Staubli VAL3: HMI_util.pjx

--- HMI_util.pjx ---
Parameters version=s8.12.2Cs9_BS2561 stackSize=5000 millimeterUnit=true
Program file=initJogMode.pgx
Program file=jogMode.pgx
Program file=loadingPage.pgx
Program file=login.pgx
Program file=setBtnColor.pgx
Program file=setframemode.pgx
Program file=setjointmode.pgx
Program file=setnullmode.pgx
Program file=settoolmode.pgx
Program file=start.pgx
Program file=stop.pgx
Data file=HMI_util.dtx
Library alias=savedata path=Disk://source/saveData/saveData.pjx

--- HMI_util.dtx ---
mdesc mNomSpeed
public string sShowType[6]
public string sShowNum[6]
public string sJoint[6]
  [0] = "J1:"
  [1] = "J2:"
  [2] = "J3:"
  [3] = "J4:"
  [4] = "J5:"
  [5] = "J6:"
public string sCartisiam[6]
  [0] = "X:"
  [1] = "Y:"
  [2] = "Z:"
  [3] = "RX:"
  [4] = "RY:"
  [5] = "RZ:"
public string sPage
string sInputPswd
bool bConfirm
bool bCancel
string sPassword = "1"
num nUsingTool

--- start.pgx ---
program start()
begin
end

--- initJogMode.pgx ---
public program initJogMode()
  local num l_i
begin
   for l_i = 0 to size(sShowType)-1
    sShowType[l_i]=sCartisiam[l_i]
  endFor
end

--- jogMode.pgx ---
public program jogMode(num x_nToolIndex, num x_nFrameIndex)
  local num l_nJogMode
  local jointRx l_jHere
  local pointRx l_pHere
  local tool l_tTool
  local frame l_fFrame
begin
  link(l_tTool,flange)
  link(l_fFrame,world)
  l_nJogMode=$getJogmode()
  l_jHere=herej()
  call savedata:getTool(x_nToolIndex,l_tTool)
  call savedata:getFrame(x_nFrameIndex,l_fFrame)
  l_pHere=here(l_tTool,l_fFrame)
  switch l_nJogMode
    case 0
      call setBtnColor(0)
      sShowNum[0]=toString(".2",l_pHere.trsf.x)
      sShowNum[1]=toString(".2",l_pHere.trsf.y)
      sShowNum[2]=toString(".2",l_pHere.trsf.z)
      sShowNum[3]=toString(".2",l_pHere.trsf.rx)
      sShowNum[4]=toString(".2",l_pHere.trsf.ry)
      sShowNum[5]=toString(".2",l_pHere.trsf.rz )
    break
    case 1
      call setBtnColor(1)
      sShowNum[0]=toString(".2",l_jHere.j1)
      sShowNum[1]=toString(".2",l_jHere.j2)
      sShowNum[2]=toString(".2",l_jHere.j3)
      sShowNum[3]=toString(".2",l_jHere.j4)
      sShowNum[4]=toString(".2",l_jHere.j5)
      sShowNum[5]=toString(".2",l_jHere.j6)
    break
    case 2
      call setBtnColor(2)
      sShowNum[0]=toString(".2",l_pHere.trsf.x)
      sShowNum[1]=toString(".2",l_pHere.trsf.y)
      sShowNum[2]=toString(".2",l_pHere.trsf.z)
      sShowNum[3]=toString(".2",l_pHere.trsf.rx)
      sShowNum[4]=toString(".2",l_pHere.trsf.ry)
      sShowNum[5]=toString(".2",l_pHere.trsf.rz )
    break
    case 3
      call setBtnColor(3)
      sShowNum[0]=toString(".2",l_pHere.trsf.x)
      sShowNum[1]=toString(".2",l_pHere.trsf.y)
      sShowNum[2]=toString(".2",l_pHere.trsf.z)
      sShowNum[3]=toString(".2",l_pHere.trsf.rx)
      sShowNum[4]=toString(".2",l_pHere.trsf.ry)
      sShowNum[5]=toString(".2",l_pHere.trsf.rz )
    break
  endSwitch
end

--- loadingPage.pgx ---
public program loadingPage()
begin
  userPage("loading")
  delay(0)
end

--- login.pgx ---
public program login(bool& x_bResult)
  local bool l_bCancel
begin
  sPage=""
  x_bResult=false
  do
    if sPage!="login"
      sPage="login"
      //init
      sInputPswd=""
      //bind
      userPageBind("login","pwd1","value",sInputPswd,1,"rw")
      userPageBindClick("login","btn1",bConfirm,true)
      userPageBindClick("login","btn2",bCancel,true)
      //
      userPage(sPage)
      delay(0.5)
    endIf
    //button
    if bConfirm
      bConfirm=false
      if sInputPswd==sPassword
        x_bResult=true
      else
        userPageAlert("invalid password!")
      endIf
    elseIf bCancel
      bCancel=false
      l_bCancel=true
    endIf




    delay(0)
  until l_bCancel==true
end

--- setBtnColor.pgx ---
public program setBtnColor(num x_nJogmode)
  local string l_sNULLcolor
  local num l_i
  local string l_sbtn
  local string l_sSELcolor
begin
  l_sNULLcolor="#FFFFFF"
  l_sSELcolor="#3399FF"

  switch x_nJogmode
    case 0
      for l_i = 1 to 4 step 1
        l_sbtn="btn"+toString("",l_i)
        userPageSet("jogmode",l_sbtn,"style.backgroundColor",l_sNULLcolor)
      endFor
    break
    case 1
      userPageSet("jogmode","btn1","style.backgroundColor",l_sNULLcolor)
      userPageSet("jogmode","btn2","style.backgroundColor",l_sSELcolor)
      userPageSet("jogmode","btn3","style.backgroundColor",l_sNULLcolor)
      userPageSet("jogmode","btn4","style.backgroundColor",l_sNULLcolor)
    break
    case 2
      userPageSet("jogmode","btn1","style.backgroundColor",l_sNULLcolor)
      userPageSet("jogmode","btn3","style.backgroundColor",l_sSELcolor)
      userPageSet("jogmode","btn2","style.backgroundColor",l_sNULLcolor)
      userPageSet("jogmode","btn4","style.backgroundColor",l_sNULLcolor)
    break
    case 3
      userPageSet("jogmode","btn1","style.backgroundColor",l_sNULLcolor)
      userPageSet("jogmode","btn2","style.backgroundColor",l_sNULLcolor)
      userPageSet("jogmode","btn3","style.backgroundColor",l_sNULLcolor)
      userPageSet("jogmode","btn4","style.backgroundColor",l_sSELcolor)
    break

  endSwitch
end

--- setframemode.pgx ---
public program setframemode()
  local num l_i
begin
  $jogMode(2)
  for l_i = 0 to size(sShowType)-1
    sShowType[l_i]=sCartisiam[l_i]
  endFor
end

--- setjointmode.pgx ---
public program setjointmode()
  local num l_i
begin
  $jogMode(1)
   for l_i = 0 to size(sShowType)-1
    sShowType[l_i]=sJoint[l_i]
  endFor
end

--- setnullmode.pgx ---
public program setnullmode()
  local num l_i
begin
  $jogMode(0)
   for l_i = 0 to size(sShowType)-1
    sShowType[l_i]=sCartisiam[l_i]
  endFor
end

--- settoolmode.pgx ---
public program settoolmode()
  local num l_i
begin
  $jogMode(3)
   for l_i = 0 to size(sShowType)-1
    sShowType[l_i]=sCartisiam[l_i]
  endFor
end

--- stop.pgx ---
program stop()
begin
end
